(* IEC 61131-3 sources: s7-to-codesys/tests/POUs/S7Compat/FB_StandardFlipFlop_Test, 5 files *)

(* ---- RsResetDominant.method.decl.st ---- *)
// RS Standard: при SET = RESET1 = TRUE выход Q1 = FALSE (сброс главнее).
METHOD PRIVATE RsResetDominant
VAR
    fbDut : RS;     // проверяемый элемент (новый экземпляр на каждый вызов метода)
END_VAR

(* ---- RsSetHeldReappliesAfterReset.method.decl.st ---- *)
// Справка Standard пишет о входах «Rising edge», модель stsim — по уровню (МЭК 61131-3). Тест различает:
// SET держится TRUE, RESET1 импульсом сбрасывает Q1; после снятия RESET1 по уровню Q1 снова TRUE,
// по фронту осталась бы FALSE.
METHOD PRIVATE RsSetHeldReappliesAfterReset
VAR
    fbDut : RS;     // проверяемый элемент (новый экземпляр на каждый вызов метода)
END_VAR

(* ---- S7RsSetDominantViaSr.method.decl.st ---- *)
// S7 RS (R, S1): «сначала R, потом S» — при R = S1 = 1 выход установлен. Перевод s7conv: CODESYS SR
// (SET1 := S1, RESET := R, Q1 — выход Q).
METHOD PRIVATE S7RsSetDominantViaSr
VAR
    fbDut : SR;     // перевод экземпляра S7 RS (новый экземпляр на каждый вызов метода)
END_VAR

(* ---- S7SrResetDominantViaRs.method.decl.st ---- *)
// S7 SR (S, R1): «сначала S, потом R» — при S = R1 = 1 выход сброшен. Перевод s7conv: CODESYS RS
// (SET := S, RESET1 := R1, Q1 — выход Q).
METHOD PRIVATE S7SrResetDominantViaRs
VAR
    fbDut : RS;     // перевод экземпляра S7 SR (новый экземпляр на каждый вызов метода)
END_VAR

(* ---- SrSetDominant.method.decl.st ---- *)
// SR Standard: при SET1 = RESET = TRUE выход Q1 = TRUE (установка главнее); вход SET1 сброшен — Q1 держится.
METHOD PRIVATE SrSetDominant
VAR
    fbDut : SR;     // проверяемый элемент (новый экземпляр на каждый вызов метода)
END_VAR
